// TIA Portal V15.1 export
// export: Created 2026-11-02T18:55:11.539963Z, ExportSetting WithDefaults, DisplayName Totally Integrated Automation Portal, DisplayVersion V15.1, DisplayName TIA Portal Openness, DisplayVersion V15.1, DisplayName STEP 7 Professional, DisplayVersion V15.1, DisplayName WinCC Professional, DisplayVersion V15.1
ORGANIZATION_BLOCK "Startup"   // OB100, LAD, Startup
TITLE = Startup
{ S7_Optimized_Access := 'TRUE' }
VERSION : 0.1
// Startup OB (decisions/0006)
// stored: AutoNumber false, IsIECCheckEnabled false, SetENOAutomatically False
   VAR_INPUT
      LostRetentive : Bool;   // True if retentive data are lost
      LostRTC : Bool;   // True if date and time are lost
   END_VAR
BEGIN

REGION Network 1: C02 — power-up: first-scan flag (scrubber trips, burners need START)
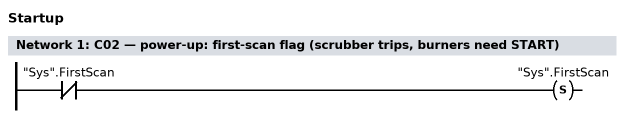
   RUNG wire#powerrail
      I_Contact( "Sys".FirstScan )
      S_Coil( "Sys".FirstScan )
   END_RUNG
   // the same network as SCL:
   IF NOT "Sys".FirstScan THEN "Sys".FirstScan := TRUE; END_IF;
END_REGION
END_ORGANIZATION_BLOCK
